(* IEC 61131-3 sources: SRCI_CLIENT_PLC/RobotLibrary/Library/POUs/Additional/MC_AvoidSingularity/Structures, 4 files *)

(* ---- AvoidSingularityOutCmd.st ---- *)
{attribute 'pack_mode' := '1'}
// -------------------------------------------------------------------------
//  SRCI Robot Library
// -------------------------------------------------------------------------
//
//  Object:      AvoidSingularityOutCmd
//  Author:      Thorsten Brach
//  Date:        2024-06-22
//
//  Description:
//
//
//  Copyright:
//    (C) 2024 Thorsten Brach. All rights reserved
//             Licensed under the MIT License.
//
//  Disclaimer:
//    This project is provided without any guarantee and can be used for
//    private and commercial purposes. Any use is at the user’s
//    own risk and responsibility.
//
// -------------------------------------------------------------------------
TYPE AvoidSingularityOutCmd :
STRUCT
END_STRUCT
END_TYPE

(* ---- AvoidSingularityParCmd.st ---- *)
{attribute 'pack_mode' := '1'}
// -------------------------------------------------------------------------
//  SRCI Robot Library
// -------------------------------------------------------------------------
//
//  Object:      AvoidSingularityParCmd
//  Author:      Thorsten Brach
//  Date:        2024-06-22
//
//  Description:
//
//
//  Copyright:
//    (C) 2024 Thorsten Brach. All rights reserved
//             Licensed under the MIT License.
//
//  Disclaimer:
//    This project is provided without any guarantee and can be used for
//    private and commercial purposes. Any use is at the user’s
//    own risk and responsibility.
//
// -------------------------------------------------------------------------
TYPE AvoidSingularityParCmd :
STRUCT
  /// Define in which way the singularity should be avoided
  Mode : SingularityAvoidanceMode;
END_STRUCT
END_TYPE

(* ---- AvoidSingularityRecvData.st ---- *)
{attribute 'pack_mode' := '1'}
// -------------------------------------------------------------------------
//  SRCI Robot Library
// -------------------------------------------------------------------------
//
//  Object:      AvoidSingularityRecvData
//  Author:      Thorsten Brach
//  Date:        2024-06-22
//
//  Description:
//
//
//  Copyright:
//    (C) 2024 Thorsten Brach. All rights reserved
//             Licensed under the MIT License.
//
//  Disclaimer:
//    This project is provided without any guarantee and can be used for
//    private and commercial purposes. Any use is at the user’s
//    own risk and responsibility.
//
// -------------------------------------------------------------------------
TYPE AvoidSingularityRecvData EXTENDS RspHeader :
STRUCT
  /// TRUE when robot is set to RA power state "Enabled".
  Enabled : BOOL;
END_STRUCT
END_TYPE

(* ---- AvoidSingularitySendData.st ---- *)
{attribute 'pack_mode' := '1'}
// -------------------------------------------------------------------------
//  SRCI Robot Library
// -------------------------------------------------------------------------
//
//  Object:      AvoidSingularitySendData
//  Author:      Thorsten Brach
//  Date:        2024-06-22
//
//  Description:
//
//
//  Copyright:
//    (C) 2024 Thorsten Brach. All rights reserved
//             Licensed under the MIT License.
//
//  Disclaimer:
//    This project is provided without any guarantee and can be used for
//    private and commercial purposes. Any use is at the user’s
//    own risk and responsibility.
//
// -------------------------------------------------------------------------
TYPE AvoidSingularitySendData EXTENDS CmdHeader:
STRUCT
  /// Set TRUE to activate avoid singularity mode
  Enable : BOOL;
  /// Define in which way the singularity should be avoided
  Mode   : SingularityAvoidanceMode;
END_STRUCT
END_TYPE
